(* PLC project , Example Feedback *)

PROGRAM Toggle
  VAR
    Q : BOOL;
    Label : STRING := 'Initial String';
  END_VAR
  VAR  (* added by the conversion: wires and edge detectors of the diagram *)
    _NOT1_OUT : BOOL;
  END_VAR

(* FBD diagram, written out as Structured Text *)
_NOT1_OUT := NOT _NOT1_OUT;
Q := _NOT1_OUT;
END_PROGRAM

CONFIGURATION c
  RESOURCE r ON PLC
    TASK t(INTERVAL := T#20ms, PRIORITY := 1);
    PROGRAM i WITH t : Toggle;
  END_RESOURCE
END_CONFIGURATION
